Fanuc KAREL source: kb00119.KL

PROGRAM KB00119
%STACKSIZE=65535
%PRIORITY=65535
%NOLOCKGROUP
VAR
P1 : INTEGER
P2 : INTEGER
BEGIN
P1=1
P2=1
LOCK_GROUP(P1,P2)
END KB00119
